(* IEC 61131-3 sources: sis-interlock-demo/src/POUs/Generated/PRG_Sis, 1 file *)

(* ---- PRG_Sis.decl.st ---- *)
// AUTO-GENERATED by cemgen 1.0.0 — не редактировать: правьте матрицу и запустите
//   python -m cemgen generate <файл матрицы .csv или .xlsx>
// Матрица: SIS-V101-CEM, объект V-101, ревизия B от 2026-10-19, SHA-256 сетки df2ed4841a9453ca
// Назначение: цикл ПАЗ объекта V-101: вызов GVL_Sis.fbApp с системным временем, журналом, образом
//             ввода-вывода и командами HMI. Вызывается из PRG_Main (MainTask).
// Автор:      kr0nsch; код — генератор cemgen
// Версия:     1.0.0
// Документ:   docs/DESIGN.md, раздел «10. Генератор cemgen»; docs/cause_effect_matrix.md
// ВНИМАНИЕ:   код демонстрационный и не предназначен для систем безопасности. Реальная ПАЗ требует
//             определения SIL, сертифицированных аппаратных и программных средств и валидации по
//             ГОСТ Р МЭК 61511.
PROGRAM PRG_Sis
VAR
END_VAR
